(* IEC 61131-3 sources: volt/packages/volt-lsp-iec/test-corpus/CodesysTestProject/Device/Plc Logic/Application/Library Manager/CmpEventMgr Implementation, 22 files *)

(* ---- EVENTCLOSE.pou ---- *)
FUNCTION EVENTCLOSE : RTS_IEC_RESULT
VAR_INPUT
	HEVENT : RTS_IEC_HANDLE;
END_VAR
VAR_IN_OUT
	RESULT : RTS_IEC_RESULT;
END_VAR
END_FUNCTION

(* ---- EVENTCLOSE2.pou ---- *)
FUNCTION EVENTCLOSE2 : RTS_IEC_RESULT
VAR_INPUT
	HEVENT : RTS_IEC_HANDLE;
END_VAR
END_FUNCTION

(* ---- EVENTCREATE.pou ---- *)
FUNCTION EVENTCREATE : RTS_IEC_HANDLE
VAR_INPUT
	EVENTID : UDINT;
	CMPIDPROVIDER : UDINT;
END_VAR
VAR_IN_OUT
	RESULT : RTS_IEC_RESULT;
END_VAR
END_FUNCTION

(* ---- EVENTCREATE2.pou ---- *)
FUNCTION EVENTCREATE2 : RTS_IEC_HANDLE
VAR_INPUT
	EVENTID : UDINT;
	CMPIDPROVIDER : UDINT;
	NCALLBACKSPOSSIBLE : UDINT;
END_VAR
VAR_IN_OUT
	RESULT : RTS_IEC_RESULT;
END_VAR
END_FUNCTION

(* ---- EVENTCREATEEVENTID.pou ---- *)
FUNCTION EVENTCREATEEVENTID : UDINT
VAR_INPUT
	EVENT : UINT;
	CLASS : UINT;
END_VAR
VAR_IN_OUT
	RESULT : RTS_IEC_RESULT;
END_VAR
END_FUNCTION

(* ---- EVENTDELETE.pou ---- *)
FUNCTION EVENTDELETE : RTS_IEC_RESULT
VAR_INPUT
	HEVENT : RTS_IEC_HANDLE;
END_VAR
VAR_IN_OUT
	RESULT : RTS_IEC_RESULT;
END_VAR
END_FUNCTION

(* ---- EVENTDELETE2.pou ---- *)
FUNCTION EVENTDELETE2 : RTS_IEC_RESULT
VAR_INPUT
	HEVENT : RTS_IEC_HANDLE;
END_VAR
END_FUNCTION

(* ---- EVENTGETCLASS.pou ---- *)
FUNCTION EVENTGETCLASS : UINT
VAR_INPUT
	EVENTID : UDINT;
END_VAR
END_FUNCTION

(* ---- EVENTGETEVENT.pou ---- *)
FUNCTION EVENTGETEVENT : UINT
VAR_INPUT
	EVENTID : UDINT;
END_VAR
END_FUNCTION

(* ---- EVENTOPEN.pou ---- *)
FUNCTION EVENTOPEN : RTS_IEC_HANDLE
VAR_INPUT
	EVENTID : UDINT;
	CMPIDPROVIDER : UDINT;
END_VAR
VAR_IN_OUT
	RESULT : RTS_IEC_RESULT;
END_VAR
END_FUNCTION

(* ---- EVENTPOST.pou ---- *)
FUNCTION EVENTPOST : RTS_IEC_RESULT
VAR_INPUT
	HEVENT : RTS_IEC_HANDLE;
	PEVENTPARAM : POINTER TO EventParam;
END_VAR
END_FUNCTION

(* ---- EVENTPOST2.pou ---- *)
FUNCTION EVENTPOST2 : RTS_IEC_RESULT
VAR_INPUT
	HEVENT : RTS_IEC_HANDLE;
	PEVENTPARAM : POINTER TO EventParam2;
END_VAR
END_FUNCTION

(* ---- EVENTPOSTBYEVENT.pou ---- *)
FUNCTION EVENTPOSTBYEVENT : RTS_IEC_RESULT
VAR_INPUT
	EVENTID : UDINT;
	CMPIDPROVIDER : UDINT;
	PEVENTPARAM : POINTER TO EventParam;
END_VAR
END_FUNCTION

(* ---- EVENTPOSTBYEVENT2.pou ---- *)
FUNCTION EVENTPOSTBYEVENT2 : RTS_IEC_RESULT
VAR_INPUT
	EVENTID : UDINT;
	CMPIDPROVIDER : UDINT;
	PEVENTPARAM : POINTER TO EventParam2;
END_VAR
END_FUNCTION

(* ---- EVENTREGISTERCALLBACK.pou ---- *)
FUNCTION EVENTREGISTERCALLBACK : RTS_IEC_HANDLE
VAR_INPUT
	HEVENT : RTS_IEC_HANDLE;
	PICALLBACK : ICmpEventCallback;
END_VAR
VAR_IN_OUT
	RESULT : RTS_IEC_RESULT;
END_VAR
END_FUNCTION

(* ---- EVENTREGISTERCALLBACK2.pou ---- *)
FUNCTION EVENTREGISTERCALLBACK2 : RTS_IEC_HANDLE
VAR_INPUT
	HEVENT : RTS_IEC_HANDLE;
	PICALLBACK : ICmpEventCallback;
	PUSERPARAMETER : POINTER TO BYTE;
END_VAR
VAR_IN_OUT
	RESULT : RTS_IEC_RESULT;
END_VAR
END_FUNCTION

(* ---- EVENTREGISTERCALLBACKFUNCTION.pou ---- *)
FUNCTION EVENTREGISTERCALLBACKFUNCTION : RTS_IEC_RESULT
VAR_INPUT
	HEVENT : RTS_IEC_HANDLE;
	PFCALLBACKFUNCTION : POINTER TO BYTE;
END_VAR
END_FUNCTION

(* ---- EVENTREGISTERCALLBACKFUNCTION2.pou ---- *)
FUNCTION EVENTREGISTERCALLBACKFUNCTION2 : RTS_IEC_RESULT
VAR_INPUT
	HEVENT : RTS_IEC_HANDLE;
	PFCALLBACKFUNCTION : POINTER TO BYTE;
	PUSERPARAMETER : POINTER TO BYTE;
END_VAR
END_FUNCTION

(* ---- EVENTREGISTEREDCALLBACKS.pou ---- *)
FUNCTION EVENTREGISTEREDCALLBACKS : UDINT
VAR_INPUT
	HEVENT : RTS_IEC_HANDLE;
END_VAR
VAR_IN_OUT
	RESULT : RTS_IEC_RESULT;
END_VAR
END_FUNCTION

(* ---- EVENTUNREGISTERCALLBACK.pou ---- *)
FUNCTION EVENTUNREGISTERCALLBACK : RTS_IEC_RESULT
VAR_INPUT
	HEVENT : RTS_IEC_HANDLE;
	HINTERFACE : RTS_IEC_HANDLE;
END_VAR
END_FUNCTION

(* ---- EVENTUNREGISTERCALLBACKFUNCTION.pou ---- *)
FUNCTION EVENTUNREGISTERCALLBACKFUNCTION : RTS_IEC_RESULT
VAR_INPUT
	HEVENT : RTS_IEC_HANDLE;
	PFCALLBACKFUNCTION : POINTER TO BYTE;
END_VAR
END_FUNCTION

(* ---- EVENTUNREGISTERCALLBACKFUNCTION2.pou ---- *)
FUNCTION EVENTUNREGISTERCALLBACKFUNCTION2 : RTS_IEC_RESULT
VAR_INPUT
	HEVENT : RTS_IEC_HANDLE;
	PFCALLBACKFUNCTION : POINTER TO BYTE;
	PUSERPARAMETER : POINTER TO BYTE;
END_VAR
END_FUNCTION
